(* IEC 61131-3 sources: POMIRTS_lab3/AS/Library/AsSem, 2 files *)

(* ---- AsSem.fun ---- *)
(********************************************************************
 * COPYRIGHT -- Bernecker + Rainer
 ********************************************************************
 * Library: AsSem
 * File: AsSem.fun
 * Author: B+R
 ********************************************************************
 * Functions and function blocks of library AsSem
 ********************************************************************)

FUNCTION_BLOCK SemCreate				(*create semaphore; asynchronous execution*)
	VAR_INPUT
		enable			: BOOL;			(*enables execution*)
		initCount		: UDINT;		(*initial value*)
		maxCount		: UDINT;		(*maximum value*)
	END_VAR

	VAR_OUTPUT
		status			: UINT;			(*execution status: ERR_OK, ERR_FUB_ENABLE_FALSE, ERR_FUB_BUSY, 0xXXXX = see help*)
		ident			: UDINT;		(*semaphore ident*)
	END_VAR

	VAR
        i_state			: UINT;			(*internal variable*)
		i_result		: UINT;			(*internal variable*)
        i_tmp			: UDINT;		(*internal variable*)
	END_VAR
END_FUNCTION_BLOCK

FUNCTION_BLOCK SemDelete				(*delete semaphore; asynchronous execution*)
	VAR_INPUT
		enable			: BOOL;			(*enables execution*)
		ident			: UDINT;		(*semaphore ident*)
	END_VAR

	VAR_OUTPUT
		status			: UINT;			(*execution status: ERR_OK, ERR_FUB_ENABLE_FALSE, ERR_FUB_BUSY, 0xXXXX = see help*)
	END_VAR

	VAR
        i_state			: UINT;			(*internal variable*)
		i_result		: UINT;			(*internal variable*)
        i_tmp			: UDINT;		(*internal variable*)
	END_VAR
END_FUNCTION_BLOCK

FUNCTION_BLOCK SemGetInfo				(*get semaphore info*)
	VAR_INPUT
		enable			: BOOL;			(*enables execution*)
		ident			: UDINT;		(*semaphore ident*)
	END_VAR

	VAR_OUTPUT
		status			: UINT;			(*execution status: 0xXXXX = see help*)
		maxCount		: UDINT;		(*maximum value*)
		curCount		: UDINT;		(*current value*)
	END_VAR

END_FUNCTION_BLOCK

FUNCTION SemAcquire : UINT				(*acquire semaphore*)
	VAR_INPUT
		ident		:UDINT;				(*semaphore ident*)
	END_VAR
END_FUNCTION

FUNCTION SemRelease : UINT				(*release semaphore*)
	VAR_INPUT
		ident		:UDINT;				(*semaphore ident*)
	END_VAR
END_FUNCTION

(* ---- AsSem.var ---- *)
(********************************************************************
 * COPYRIGHT -- Bernecker + Rainer
 ********************************************************************
 * Library: AsSem
 * File: AsSem.var
 * Author: B+R
 ********************************************************************
 * Local variables of library AsSem
 ********************************************************************)

VAR CONSTANT
	semERR_CREATE						: UINT := 33320;	(*create semaphore error*)
	semERR_DELETE						: UINT := 33321;	(*delete semaphore error*)
	semERR_NOT_EXIST					: UINT := 33322;	(*invalid semaphore ident, check parameter*)
	semERR_NOT_FREE						: UINT := 33323;	(*semaphore already acquired*)
	semERR_ALREADY_FREE					: UINT := 33324;	(*semaphore not acquired*)
END_VAR
